          [0]
            bool bSafePoint
            ifItem iIfItem
              [0]
                bool bANDOR[2]
                num nSigIndex[3]
                num nSigType[3]
                num nValue[3]
            mdesc mMdesc
            num nActionIndex = 42
            num nDelay
            num nMoveType = 1
            num nPercentage
            num nSigValue = 1
        pointRx pPointRx[2] = {x=-245.0810672, y=-321.451661, z=639.817242, rx=-2.232299, ry=1.28487, rz=0.967617, shoulder=lefty, elbow=enegative, wrist=wpositive}
        string sID
      [8]
        bool bMarked
        jointRx jJointRx = {j1=-122.510061, j2=129.763772, j3=-115.645271, j4=180.40219, j5=16.691098, j6=-56.935013}
        pointRx pInter
        paraItem pParaItem
          [0]
            bool bSafePoint
            ifItem iIfItem
              [0]
                bool bANDOR[2]
                num nSigIndex[3]
                num nSigType[3]
                num nValue[3]
            mdesc mMdesc
            num nActionIndex = 42
            num nDelay
            num nMoveType = 1
            num nPercentage
            num nSigValue = 1
        pointRx pPointRx[2] = {x=-204.794752, y=-412.495541, z=639.817259, rx=-2.23161, ry=1.284656, rz=0.967787, shoulder=lefty, elbow=enegative, wrist=wpositive}
        string sID
      [9]
        bool bMarked
        jointRx jJointRx = {j1=-115.509708, j2=123.384757, j3=-95.0786351, j4=179.613978, j5=30.87235, j6=-63.211859}
        pointRx pInter
        paraItem pParaItem
          [0]
            bool bSafePoint
            ifItem iIfItem
              [0]
                bool bANDOR[2]
                num nSigIndex[3]
                num nSigType[3]
                num nValue[3]
            mdesc mMdesc
            num nActionIndex = 42
            num nDelay
            num nMoveType = 1
            num nPercentage
            num nSigValue = 1
        pointRx pPointRx[2] = {x=-204.829932, y=-549.361149, z=639.817236, rx=-2.230566, ry=1.283434, rz=0.967655, shoulder=lefty, elbow=enegative, wrist=wpositive}
        string sID
      [10]
        bool bMarked
        jointRx jJointRx = {j1=-115.168839, j2=115.765951, j3=-75.660997, j4=179.549971, j5=42.662693, j6=-65.612389}
        pointRx pInter
        paraItem pParaItem
          [0]
            bool bSafePoint
            ifItem iIfItem
              [0]
                bool bANDOR[2]
                num nSigIndex[3]
                num nSigType[3]
                num nValue[3]
            mdesc mMdesc
            num nActionIndex = 42
            num nDelay
            num nMoveType = 1
            num nPercentage
            num nSigValue = 1
        pointRx pPointRx[2] = {x=-243.328707, y=-641.656144, z=639.817272, rx=-2.184752, ry=1.363169, rz=-1.0929741, shoulder=lefty, elbow=enegative, wrist=wpositive}
        string sID
      [11]
        bool bMarked
        jointRx jJointRx = {j1=-103.18234, j2=119.0666826, j3=-83.752693, j4=178.724024, j5=37.773968, j6=-75.789236}
        pointRx pInter
        paraItem pParaItem
          [0]
            bool bSafePoint
            ifItem iIfItem
              [0]
                bool bANDOR[2]
                num nSigIndex[3]
                num nSigType[3]
                num nValue[3]
            mdesc mMdesc
            num nActionIndex = 42
            num nDelay
            num nMoveType = 1
            num nPercentage
            num nSigValue = 1
        pointRx pPointRx[2] = {x=-91.940597, y=-641.690605, z=639.817264, rx=-2.210413, ry=1.320263, rz=0.0285249, shoulder=lefty, elbow=enegative, wrist=wpositive}
        string sID
      [12]
        bool bMarked
        jointRx jJointRx = {j1=-96.605755, j2=119.651273, j3=-85.228552, j4=178.232883, j5=36.783421, j6=-81.95314}
        pointRx pInter
        paraItem pParaItem
          [0]
            bool bSafePoint
            ifItem iIfItem
              [0]
                bool bANDOR[2]
                num nSigIndex[3]
                num nSigType[3]
                num nValue[3]
            mdesc mMdesc
            num nActionIndex = 42
            num nDelay
            num nMoveType = 1
            num nPercentage
            num nSigValue = 1
        pointRx pPointRx[2] = {x=-14.68309, y=-641.690595, z=639.817262, rx=-2.210425, ry=1.321003, rz=0.029458, shoulder=lefty, elbow=enegative, wrist=wpositive}
        string sID
      [13]
        bool bMarked
        jointRx jJointRx = {j1=-101.415655, j2=125.744666, j3=-101.857376, j4=178.0690532, j5=26.328772, j6=-76.831785}
        pointRx pInter
        paraItem pParaItem
          [0]
            bool bSafePoint
            ifItem iIfItem
              [0]
                bool bANDOR[2]
                num nSigIndex[3]
                num nSigType[3]
                num nValue[3]
            mdesc mMdesc
            num nActionIndex = 42
            num nDelay
            num nMoveType = 1
            num nPercentage
            num nSigValue = 1
        pointRx pPointRx[2] = {x=-51.703517, y=-546.433248, z=639.817258, rx=-2.211187, ry=1.319905, rz=0.0291157, shoulder=lefty, elbow=enegative, wrist=wpositive}
        string sID
      [14]
        bool bMarked
        jointRx jJointRx = {j1=-104.908394, j2=131.188615, j3=-122.570612, j4=176.33465, j5=11.11624, j6=-71.475976}
        pointRx pInter
        paraItem pParaItem
          [0]
            bool bSafePoint
            ifItem iIfItem
              [0]
                bool bANDOR[2]
                num nSigIndex[3]
                num nSigType[3]
                num nValue[3]
            mdesc mMdesc
            num nActionIndex = 42
            num nDelay
            num nMoveType = 1
            num nPercentage
            num nSigValue = 1
        pointRx pPointRx[2] = {x=-51.703514, y=-412.500595, z=639.817231, rx=-2.211237, ry=1.319324, rz=0.0290677, shoulder=lefty, elbow=enegative, wrist=wpositive}
        string sID
      [15]
        bool bMarked
        jointRx jJointRx = {j1=-113.792229, j2=132.0385925, j3=-133.203423, j4=167.238796, j5=1.425916, j6=-53.439675}
        pointRx pInter
        paraItem pParaItem
          [0]
            bool bSafePoint
            ifItem iIfItem
              [0]
                bool bANDOR[2]
                num nSigIndex[3]
                num nSigType[3]
                num nValue[3]
            mdesc mMdesc
            num nActionIndex = 42
            num nDelay
            num nMoveType = 1
            num nPercentage
            num nSigValue = 1
        pointRx pPointRx[2] = {x=-86.764293, y=-327.545777, z=639.814183, rx=-2.211628, ry=1.318889, rz=0.029149, shoulder=lefty, elbow=enegative, wrist=wpositive}
        string sID
      [16]
        bool bMarked
        jointRx jJointRx = {j1=-111.801102, j2=131.0492813, j3=-121.763212, j4=165.182491, j5=10.00939302, j6=-125.703677}
        pointRx pInter
        paraItem pParaItem
          [0]
            bool bSafePoint
            ifItem iIfItem
              [0]
                bool bANDOR[2]
                num nSigIndex[3]
                num nSigType[3]
                num nValue[3]
            mdesc mMdesc
            num nActionIndex = 42
            num nDelay
            num nMoveType = 1
            num nPercentage
            num nSigValue = 1
        pointRx pPointRx[2] = {x=-94.727754, y=-431.297828, z=639.823313, rx=0.578297, ry=2.512713, rz=-72.12797, shoulder=lefty, elbow=enegative, wrist=wpositive}
        string sID
      [17]
        bool bMarked
        jointRx jJointRx = {j1=-100.696291, j2=131.394596, j3=-123.887641, j4=160.749292, j5=7.838779, j6=-132.328285}
        pointRx pInter
        paraItem pParaItem
          [0]
            bool bSafePoint
            ifItem iIfItem
              [0]
                bool bANDOR[2]
                num nSigIndex[3]
                num nSigType[3]
                num nValue[3]
            mdesc mMdesc
            num nActionIndex = 42
            num nDelay
            num nMoveType = 1
            num nPercentage
            num nSigValue = 1
        pointRx pPointRx[2] = {x=-7.700551, y=-431.29776, z=639.823315, rx=0.578366, ry=2.513634, rz=-72.118873, shoulder=lefty, elbow=enegative, wrist=wpositive}
        string sID
      [18]
        bool bMarked
        jointRx jJointRx = {j1=-85.175274, j2=131.219929, j3=-122.767363, j4=172.20701, j5=10.687341, j6=-85.487938}
        pointRx pInter
        paraItem pParaItem
          [0]
            bool bSafePoint
            ifItem iIfItem
              [0]
                bool bANDOR[2]
                num nSigIndex[3]
                num nSigType[3]
                num nValue[3]
            mdesc mMdesc
            num nActionIndex = 42
            num nDelay
            num nMoveType = 1
            num nPercentage
            num nSigValue = 1
        pointRx pPointRx[2] = {x=97.129831, y=-406.771802, z=639.823216, rx=-2.251869, ry=1.255999, rz=1.675152, shoulder=lefty, elbow=enegative, wrist=wpositive}
        string sID
      [19]
        bool bMarked
        jointRx jJointRx = {j1=-78.327634, j2=132.0275027, j3=-133.511556, j4=105.524405, j5=1.749155, j6=-25.524463}
        pointRx pInter
        paraItem pParaItem
          [0]
            bool bSafePoint
            ifItem iIfItem
              [0]
                bool bANDOR[2]
                num nSigIndex[3]
                num nSigType[3]
                num nValue[3]
            mdesc mMdesc
            num nActionIndex = 42
            num nDelay
            num nMoveType
            num nPercentage
            num nSigValue = 1
        pointRx pPointRx[2] = {x=131.681956, y=-317.592689, z=639.818955, rx=-2.252815, ry=1.25559, rz=1.675166, shoulder=lefty, elbow=enegative, wrist=wpositive}
        string sID
      [20]
        bool bMarked
        jointRx jJointRx = {j1=-86.344906, j2=125.635703, j3=-101.533058, j4=176.84641, j5=26.303372, j6=-89.150638}
        pointRx pInter
        paraItem pParaItem
          [0]
            bool bSafePoint
            ifItem iIfItem
              [0]
                bool bANDOR[2]
                num nSigIndex[3]
                num nSigType[3]
                num nValue[3]
            mdesc mMdesc
            num nActionIndex = 42
            num nDelay
            num nMoveType = 1
            num nPercentage
            num nSigValue = 1
        pointRx pPointRx[2] = {x=97.129791, y=-544.994507, z=639.823164, rx=-2.250847, ry=1.25596, rz=1.67509, shoulder=lefty, elbow=enegative, wrist=wpositive}
        string sID
      [21]
        bool bMarked
        jointRx jJointRx = {j1=-90.472886, j2=120.653514, j3=-87.796909, j4=177.850277, j5=35.136858, j6=-86.0941041}
        pointRx pInter
        paraItem pParaItem
          [0]
            bool bSafePoint
            ifItem iIfItem
              [0]
                bool bANDOR[2]
                num nSigIndex[3]
                num nSigType[3]
                num nValue[3]
            mdesc mMdesc
            num nActionIndex = 42
            num nDelay
            num nMoveType = 1
            num nPercentage
            num nSigValue = 1
        pointRx pPointRx[2] = {x=55.621844, y=-626.948778, z=639.823217, rx=-2.25099, ry=1.255655, rz=1.674992, shoulder=lefty, elbow=enegative, wrist=wpositive}
        string sID
      [22]
        bool bMarked
        jointRx jJointRx = {j1=-83.248503, j2=126.765701, j3=-105.0119337, j4=185.0332952, j5=23.463189, j6=-12.861735}
        pointRx pInter
        paraItem pParaItem
          [0]
            bool bSafePoint
            ifItem iIfItem
              [0]
                bool bANDOR[2]
                num nSigIndex[3]
                num nSigType[3]
                num nValue[3]
            mdesc mMdesc
            num nActionIndex = 42
            num nDelay
            num nMoveType = 1
            num nPercentage
            num nSigValue = 1
        pointRx pPointRx[2] = {x=95.0604108, y=-526.24744, z=639.845413, rx=-1.382011, ry=-2.179455, rz=88.510933, shoulder=lefty, elbow=enegative, wrist=wpositive}
        string sID
      [23]
        bool bMarked
        jointRx jJointRx = {j1=-102.947247, j2=123.371825, j3=-104.720974, j4=140.865912, j5=30.580144, j6=47.745938}
        pointRx pInter
        paraItem pParaItem
          [0]
            bool bSafePoint
            ifItem iIfItem
              [0]
                bool bANDOR[2]
                num nSigIndex[3]
                num nSigType[3]
                num nValue[3]
            mdesc mMdesc
            num nActionIndex = 42
            num nDelay
            num nMoveType = 1
            num nPercentage
            num nSigValue = 1
        pointRx pPointRx[2] = {x=95.0560257, y=-526.230668, z=639.854281, rx=-1.467206, ry=19.573094, rz=89.0544323, shoulder=lefty, elbow=enegative, wrist=wpositive}
        string sID
      [24]
        bool bMarked
        jointRx jJointRx = {j1=-105.42444, j2=126.319202, j3=-118.0699052, j4=127.900909, j5=23.640583, j6=64.972841}
        pointRx pInter
        paraItem pParaItem
          [0]
            bool bSafePoint
            ifItem iIfItem
              [0]
                bool bANDOR[2]
                num nSigIndex[3]
                num nSigType[3]
                num nValue[3]
            mdesc mMdesc
            num nActionIndex = 42
            num nDelay
            num nMoveType = 1
            num nPercentage
            num nSigValue = 1
        pointRx pPointRx[2] = {x=95.0558629, y=-438.311234, z=639.854334, rx=-1.468101, ry=19.566479, rz=89.0544973, shoulder=lefty, elbow=enegative, wrist=wpositive}
        string sID
      [25]
        bool bMarked
        jointRx jJointRx = {j1=-112.0262192, j2=125.853254, j3=-136.407591, j4=84.864182, j5=17.615577, j6=117.594482}
        pointRx pInter
        paraItem pParaItem
          [0]
            bool bSafePoint
            ifItem iIfItem
              [0]
                bool bANDOR[2]
                num nSigIndex[3]
                num nSigType[3]
                num nValue[3]
            mdesc mMdesc
            num nActionIndex = 42
            num nDelay
            num nMoveType = 1
            num nPercentage
            num nSigValue = 1
        pointRx pPointRx[2] = {x=95.0562279, y=-300.211931, z=639.855152, rx=-1.466155, ry=19.566406, rz=89.0540412, shoulder=lefty, elbow=enegative, wrist=wpositive}
        string sID
      [26]
        bool bMarked
        jointRx jJointRx = {j1=-98.853409, j2=130.526556, j3=-129.84131, j4=190.937055, j5=1.850619, j6=112.778311}
        pointRx pInter
        paraItem pParaItem
          [0]
            bool bSafePoint
            ifItem iIfItem
              [0]
                bool bANDOR[2]
                num nSigIndex[3]
                num nSigType[3]
                num nValue[3]
            mdesc mMdesc
            num nActionIndex = 42
            num nDelay
            num nMoveType = 1
            num nPercentage
            num nSigValue = 1
        pointRx pPointRx[2] = {x=-10.299262, y=-371.0877835, z=648.6975, rx=-1.172321, ry=-0.172701, rz=-155.141909, shoulder=lefty, elbow=enegative, wrist=wpositive}
        string sID
      [27]
        bool bMarked
        jointRx jJointRx = {j1=-87.556691, j2=130.508226, j3=-129.0706324, j4=182.704505, j5=2.618876, j6=109.713672}
        pointRx pInter
        paraItem pParaItem
          [0]
            bool bSafePoint
            ifItem iIfItem
              [0]
                bool bANDOR[2]
                num nSigIndex[3]
                num nSigType[3]
                num nValue[3]
            mdesc mMdesc
            num nActionIndex = 42
            num nDelay
            num nMoveType = 1
            num nPercentage
            num nSigValue = 1
        pointRx pPointRx[2] = {x=64.800708, y=-371.087733, z=648.697509, rx=-1.172034, ry=-0.173648, rz=-155.14184, shoulder=lefty, elbow=enegative, wrist=wpositive}
        string sID
      [28]
        bool bMarked
        jointRx jJointRx = {j1=-76.56227, j2=130.441663, j3=-127.63649, j4=178.503737, j5=3.987538, j6=102.915897}
        pointRx pInter
        paraItem pParaItem
          [0]
            bool bSafePoint
            ifItem iIfItem
              [0]
                bool bANDOR[2]
                num nSigIndex[3]
                num nSigType[3]
                num nValue[3]
            mdesc mMdesc
            num nActionIndex = 42
            num nDelay
            num nMoveType = 1
            num nPercentage
            num nSigValue = 1
        pointRx pPointRx[2] = {x=138.739125, y=-361.605648, z=648.697463, rx=-1.172859, ry=-0.173244, rz=-155.141862, shoulder=lefty, elbow=enegative, wrist=wpositive}
        string sID
      [29]
        bool bMarked
        jointRx jJointRx = {j1=-65.258595, j2=131.722388, j3=-131.258412, j4=149.998176, j5=1.563572, j6=95.282187}
        pointRx pInter
        paraItem pParaItem
          [0]
            bool bSafePoint
            ifItem iIfItem
              [0]
                bool bANDOR[2]
                num nSigIndex[3]
                num nSigType[3]
                num nValue[3]
            mdesc mMdesc
            num nActionIndex = 42
            num nDelay
            num nMoveType = 1
            num nPercentage
            num nSigValue = 1
        pointRx pPointRx[2] = {x=203.481922, y=-305.793086, z=642.0323173, rx=-1.135624, ry=0.337465, rz=-179.971722, shoulder=lefty, elbow=enegative, wrist=wpositive}
        string sID
      [30]
        bool bMarked
        jointRx jJointRx = {j1=-75.287181, j2=130.366871, j3=-119.512671, j4=177.0231421, j5=11.88329, j6=78.230615}
        pointRx pInter
        paraItem pParaItem
          [0]
            bool bSafePoint
            ifItem iIfItem
              [0]
                bool bANDOR[2]
                num nSigIndex[3]
                num nSigType[3]
                num nValue[3]
            mdesc mMdesc
            num nActionIndex = 42
            num nDelay
            num nMoveType = 1
            num nPercentage
            num nSigValue = 1
        pointRx pPointRx[2] = {x=166.551107, y=-416.353492, z=642.0259775, rx=-1.135878, ry=0.33525, rz=-179.971835, shoulder=lefty, elbow=enegative, wrist=wpositive}
        string sID
      [31]
        bool bMarked
        jointRx jJointRx = {j1=-78.750875, j2=124.345332, j3=-98.32121, j4=178.789895, j5=27.0774003, j6=79.858309}
        pointRx pInter
        paraItem pParaItem
          [0]
            bool bSafePoint
            ifItem iIfItem
              [0]
                bool bANDOR[2]
                num nSigIndex[3]
                num nSigType[3]
                num nValue[3]
            mdesc mMdesc
            num nActionIndex = 42
            num nDelay
            num nMoveType = 1
            num nPercentage
            num nSigValue = 1
        pointRx pPointRx[2] = {x=166.551118, y=-556.425136, z=642.0259681, rx=-1.135398, ry=0.335774, rz=-179.971779, shoulder=lefty, elbow=enegative, wrist=wpositive}
        string sID
      [32]
        bool bMarked
        jointRx jJointRx = {j1=-83.872725, j2=117.4103, j3=-80.0479523, j4=179.268733, j5=38.458687, j6=84.472525}
        pointRx pInter
        paraItem pParaItem
          [0]
            bool bSafePoint
            ifItem iIfItem
              [0]
                bool bANDOR[2]
                num nSigIndex[3]
                num nSigType[3]
                num nValue[3]
            mdesc mMdesc
            num nActionIndex = 42
            num nDelay
            num nMoveType = 1
            num nPercentage
            num nSigValue = 1
        pointRx pPointRx[2] = {x=125.777964, y=-666.0321845, z=642.0361412, rx=-1.136355, ry=0.335436, rz=-179.973852, shoulder=lefty, elbow=enegative, wrist=wpositive}
        string sID
      [33]
        bool bMarked
        jointRx jJointRx = {j1=-78.0158878, j2=116.00480506, j3=-76.619863, j4=179.128646, j5=40.428713, j6=78.707523}
        pointRx pInter
        paraItem pParaItem
          [0]
            bool bSafePoint
            ifItem iIfItem
              [0]
                bool bANDOR[2]
                num nSigIndex[3]
                num nSigType[3]
                num nValue[3]
            mdesc mMdesc
            num nActionIndex = 42
            num nDelay
            num nMoveType = 1
            num nPercentage
            num nSigValue = 1
        pointRx pPointRx[2] = {x=197.538696, y=-666.0666154, z=642.0361247, rx=-1.135138, ry=0.336712, rz=-179.973468, shoulder=lefty, elbow=enegative, wrist=wpositive}
        string sID
      [34]
        bool bMarked
        jointRx jJointRx = {j1=-72.0822941, j2=113.707363, j3=-71.14889, j4=179.0271553, j5=43.540761, j6=72.816847}
        pointRx pInter
        paraItem pParaItem
          [0]
            bool bSafePoint
            ifItem iIfItem
              [0]
                bool bANDOR[2]
                num nSigIndex[3]
                num nSigType[3]
                num nValue[3]
            mdesc mMdesc
            num nActionIndex = 42
            num nDelay
            num nMoveType = 1
            num nPercentage
            num nSigValue = 1
        pointRx pPointRx[2] = {x=274.0463743, y=-666.0377191, z=642.0648113, rx=-1.136874, ry=0.336734, rz=-179.973059, shoulder=lefty, elbow=enegative, wrist=wpositive}
        string sID
      [35]
        bool bMarked
        jointRx jJointRx = {j1=-68.231832, j2=114.0101375, j3=-71.862732, j4=178.925387, j5=43.085151, j6=69.0461931}
        pointRx pInter
        paraItem pParaItem
          [0]
            bool bSafePoint
            ifItem iIfItem
              [0]
                bool bANDOR[2]
                num nSigIndex[3]
                num nSigType[3]
                num nValue[3]
            mdesc mMdesc
            num nActionIndex = 42
            num nDelay
            num nMoveType = 1
            num nPercentage
            num nSigValue = 1
        pointRx pPointRx[2] = {x=317.646205, y=-643.356636, z=642.0648372, rx=-1.138401, ry=0.335813, rz=-179.973153, shoulder=lefty, elbow=enegative, wrist=wpositive}
        string sID
      [36]
        bool bMarked
        jointRx jJointRx = {j1=-65.210051, j2=120.724606, j3=-88.443145, j4=178.570875, j5=33.182263, j6=66.435792}
        pointRx pInter
        paraItem pParaItem
          [0]
            bool bSafePoint
            ifItem iIfItem
              [0]
                bool bANDOR[2]
                num nSigIndex[3]
                num nSigType[3]
                num nValue[3]
            mdesc mMdesc
            num nActionIndex = 42
            num nDelay
            num nMoveType = 1
            num nPercentage
            num nSigValue = 1
        pointRx pPointRx[2] = {x=317.646188, y=-552.240414, z=642.0648293, rx=-1.138291, ry=0.335792, rz=-179.973173, shoulder=lefty, elbow=enegative, wrist=wpositive}
        string sID
      [37]
        bool bMarked
        jointRx jJointRx = {j1=-59.269672, j2=127.333625, j3=-107.550013, j4=177.526605, j5=20.607904, j6=61.614613}
        pointRx pInter
        paraItem pParaItem
          [0]
            bool bSafePoint
            ifItem iIfItem
              [0]
                bool bANDOR[2]
                num nSigIndex[3]
                num nSigType[3]
                num nValue[3]
            mdesc mMdesc
            num nActionIndex = 42
            num nDelay
            num nMoveType = 1
            num nPercentage
            num nSigValue = 1
        pointRx pPointRx[2] = {x=317.646169, y=-421.622338, z=642.0648205, rx=-1.138138, ry=0.335927, rz=-179.973153, shoulder=lefty, elbow=enegative, wrist=wpositive}
        string sID
      [38]
        bool bMarked
        jointRx jJointRx = {j1=-56.529834, j2=131.219574, j3=-124.66737, j4=172.915754, j5=7.371604, j6=63.585523}
        pointRx pInter
        paraItem pParaItem
          [0]
            bool bSafePoint
            ifItem iIfItem
              [0]
                bool bANDOR[2]
                num nSigIndex[3]
                num nSigType[3]
                num nValue[3]
            mdesc mMdesc
            num nActionIndex = 42
            num nDelay
            num nMoveType = 1
            num nPercentage
            num nSigValue = 1
        pointRx pPointRx[2] = {x=275.258961, y=-311.334534, z=642.0647626, rx=-1.137088, ry=0.335146, rz=-179.97331, shoulder=lefty, elbow=enegative, wrist=wpositive}
        string sID
      [39]
        bool bMarked
        jointRx jJointRx = {j1=-63.306074, j2=128.457716, j3=-111.487898, j4=177.354165, j5=17.85182, j6=65.854127}
        pointRx pInter
        paraItem pParaItem
          [0]
            bool bSafePoint
            ifItem iIfItem
              [0]
                bool bANDOR[2]
                num nSigIndex[3]
                num nSigType[3]
                num nValue[3]
            mdesc mMdesc
            num nActionIndex = 42
            num nDelay
            num nMoveType = 1
            num nPercentage
            num nSigValue = 1
        pointRx pPointRx[2] = {x=275.293372, y=-420.450747, z=642.0648054, rx=-1.136295, ry=0.336239, rz=-179.973341, shoulder=lefty, elbow=enegative, wrist=wpositive}
        string sID
      [40]
        bool bMarked
        jointRx jJointRx = {j1=-81.00112581, j2=130.644686, j3=-121.00772478, j4=177.263665, j5=10.719901, j6=83.717831}
        pointRx pInter
        paraItem pParaItem
          [0]
            bool bSafePoint
            ifItem iIfItem
              [0]
                bool bANDOR[2]
                num nSigIndex[3]
                num nSigType[3]
                num nValue[3]
            mdesc mMdesc
            num nActionIndex = 42
            num nDelay
            num nMoveType = 1
            num nPercentage
            num nSigValue = 1
        pointRx pPointRx[2] = {x=121.697258, y=-420.415642, z=642.064816, rx=-1.13739, ry=0.335022, rz=-179.973377, shoulder=lefty, elbow=enegative, wrist=wpositive}
        string sID
      [41]
        bool bMarked
        jointRx jJointRx = {j1=-101.57564, j2=130.996968, j3=-123.11763, j4=179.378674, j5=9.0641696, j6=102.209948}
        pointRx pInter
        paraItem pParaItem
          [0]
            bool bSafePoint
            ifItem iIfItem
              [0]
                bool bANDOR[2]
                num nSigIndex[3]
                num nSigType[3]
                num nValue[3]
            mdesc mMdesc
            num nActionIndex = 42
            num nDelay
            num nMoveType = 1
            num nPercentage
            num nSigValue = 1
        pointRx pPointRx[2] = {x=-34.195927, y=-420.382673, z=642.0719086, rx=-1.140588, ry=0.333521, rz=-179.976951, shoulder=lefty, elbow=enegative, wrist=wpositive}
        string sID
      [42]
        bool bMarked
        jointRx jJointRx = {j1=-117.910926, j2=130.159863, j3=-118.527747, j4=181.0779949, j5=12.798502, j6=116.877037}
        pointRx pInter
        paraItem pParaItem
          [0]
            bool bSafePoint
            ifItem iIfItem
              [0]
                bool bANDOR[2]
                num nSigIndex[3]
                num nSigType[3]
                num nValue[3]
            mdesc mMdesc
            num nActionIndex = 42
            num nDelay
            num nMoveType = 1
            num nPercentage
            num nSigValue = 1
        pointRx pPointRx[2] = {x=-168.460127, y=-420.382669, z=642.071906, rx=-1.140562, ry=0.333907, rz=-179.976921, shoulder=lefty, elbow=enegative, wrist=wpositive}
        string sID
      [43]
        bool bMarked
        jointRx jJointRx = {j1=-132.269491, j2=127.123938, j3=-106.855674, j4=181.429188, j5=21.342688, j6=130.953129}
        pointRx pInter
        paraItem pParaItem
          [0]
            bool bSafePoint
            ifItem iIfItem
              [0]
                bool bANDOR[2]
                num nSigIndex[3]
                num nSigType[3]
                num nValue[3]
            mdesc mMdesc
            num nActionIndex = 42
            num nDelay
            num nMoveType = 1
            num nPercentage
            num nSigValue = 1
        pointRx pPointRx[2] = {x=-320.674662, y=-420.382638, z=642.0718966, rx=-1.140431, ry=0.333681, rz=-179.976981, shoulder=lefty, elbow=enegative, wrist=wpositive}
        string sID
      [44]
        bool bMarked
        jointRx jJointRx = {j1=-142.441106, j2=120.824327, j3=-88.705493, j4=181.282913, j5=33.0850501, j6=141.380041}
        pointRx pInter
        paraItem pParaItem
          [0]
            bool bSafePoint
            ifItem iIfItem
              [0]
                bool bANDOR[2]
                num nSigIndex[3]
                num nSigType[3]
                num nValue[3]
            mdesc mMdesc
            num nActionIndex = 42
            num nDelay
            num nMoveType = 1
            num nPercentage
            num nSigValue = 1
        pointRx pPointRx[2] = {x=-474.689621, y=-420.382631, z=642.0718894, rx=-1.140119, ry=0.333784, rz=-179.976923, shoulder=lefty, elbow=enegative, wrist=wpositive}
        string sID
      [45]
        bool bMarked
        jointRx jJointRx = {j1=-138.108258, j2=121.207146, j3=-89.710766, j4=181.162609, j5=32.51161, j6=137.142341}
        pointRx pInter
        paraItem pParaItem
          [0]
            bool bSafePoint
            ifItem iIfItem
              [0]
                bool bANDOR[2]
                num nSigIndex[3]
                num nSigType[3]
                num nValue[3]
            mdesc mMdesc
            num nActionIndex = 42
            num nDelay
            num nMoveType = 1
            num nPercentage
            num nSigValue = 1
        pointRx pPointRx[2] = {x=-436.796862, y=-451.644484, z=642.07189, rx=-1.139469, ry=0.334472, rz=-179.976638, shoulder=lefty, elbow=enegative, wrist=wpositive}
        string sID
      [46]
        bool bMarked
        jointRx jJointRx = {j1=-127.70596, j2=126.693595, j3=-105.454305, j4=181.135682, j5=22.350888, j6=126.671469}
        pointRx pInter
        paraItem pParaItem
          [0]
            bool bSafePoint
            ifItem iIfItem
              [0]
                bool bANDOR[2]
                num nSigIndex[3]
                num nSigType[3]
                num nValue[3]
            mdesc mMdesc
            num nActionIndex = 42
            num nDelay
            num nMoveType = 1
            num nPercentage
            num nSigValue = 1
        pointRx pPointRx[2] = {x=-290.683508, y=-451.609469, z=642.07191, rx=-1.140457, ry=0.335724, rz=-179.976594, shoulder=lefty, elbow=enegative, wrist=wpositive}
        string sID
      [47]
        bool bMarked
        jointRx jJointRx = {j1=-77.238254, j2=129.340507, j3=-114.913945, j4=177.831104, j5=15.475362, j6=79.35375}
        pointRx pInter
        paraItem pParaItem
          [0]
            bool bSafePoint
            ifItem iIfItem
              [0]
                bool bANDOR[2]
                num nSigIndex[3]
                num nSigType[3]
                num nValue[3]
            mdesc mMdesc
            num nActionIndex = 42
            num nDelay
            num nMoveType = 1
            num nPercentage
            num nSigValue = 1
        pointRx pPointRx[2] = {x=158.729452, y=-451.609464, z=642.0719065, rx=-1.140389, ry=0.334964, rz=-179.976748, shoulder=lefty, elbow=enegative, wrist=wpositive}
        string sID
      [48]
        bool bMarked
        jointRx jJointRx = {j1=-63.488687, j2=124.208026, j3=-97.940675, j4=178.228458, j5=27.14867, j6=65.0910716}
        pointRx pInter
        paraItem pParaItem
          [0]
            bool bSafePoint
            ifItem iIfItem
              [0]
                bool bANDOR[2]
                num nSigIndex[3]
                num nSigType[3]
                num nValue[3]
            mdesc mMdesc
            num nActionIndex = 42
            num nDelay
            num nMoveType = 1
            num nPercentage
            num nSigValue = 1
        pointRx pPointRx[2] = {x=310.830797, y=-495.30753, z=642.0718875, rx=-1.139453, ry=0.33486, rz=-179.976891, shoulder=lefty, elbow=enegative, wrist=wpositive}
        string sID
      [49]
        bool bMarked
        jointRx jJointRx = {j1=-78.0579912, j2=127.559769, j3=-108.316642, j4=178.378161, j5=20.297351, j6=79.604006}
        pointRx pInter
        paraItem pParaItem
          [0]
            bool bSafePoint
            ifItem iIfItem
              [0]
                bool bANDOR[2]
                num nSigIndex[3]
                num nSigType[3]
                num nValue[3]
            mdesc mMdesc
            num nActionIndex = 42
            num nDelay
            num nMoveType = 1
            num nPercentage
            num nSigValue = 1
        pointRx pPointRx[2] = {x=160.873249, y=-495.272541, z=642.0719096, rx=-1.140489, ry=0.333782, rz=-179.976981, shoulder=lefty, elbow=enegative, wrist=wpositive}
        string sID
      [50]
        bool bMarked
        jointRx jJointRx = {j1=-83.970136, j2=129.00855342, j3=-113.590578, j4=181.751291, j5=14.32041, j6=-96.622719}
        pointRx pInter
        paraItem pParaItem
          [0]
            bool bSafePoint
            ifItem iIfItem
              [0]
                bool bANDOR[2]
                num nSigIndex[3]
                num nSigType[3]
                num nValue[3]
            mdesc mMdesc
            num nActionIndex = 42
            num nDelay
            num nMoveType = 1
            num nPercentage
            num nSigValue = 1
        pointRx pPointRx[2] = {x=98.789636, y=-495.232609, z=642.0875542, rx=1.143362, ry=-0.31475, rz=1.103019, shoulder=lefty, elbow=enegative, wrist=wpositive}
        string sID
      [51]
        bool bMarked
        jointRx jJointRx = {j1=-101.251443, j2=129.329307, j3=-114.876217, j4=180.377122, j5=13.270505, j6=-78.0149862}
        pointRx pInter
        paraItem pParaItem
          [0]
            bool bSafePoint
            ifItem iIfItem
              [0]
                bool bANDOR[2]
                num nSigIndex[3]
                num nSigType[3]
                num nValue[3]
            mdesc mMdesc
            num nActionIndex = 42
            num nDelay
            num nMoveType = 1
            num nPercentage
            num nSigValue = 1
        pointRx pPointRx[2] = {x=-48.311282, y=-495.232554, z=642.0875543, rx=1.143247, ry=-0.315683, rz=1.102879, shoulder=lefty, elbow=enegative, wrist=wpositive}
        string sID
      [52]
        bool bMarked
        jointRx jJointRx = {j1=-117.974593, j2=127.746571, j3=-108.963712, j4=179.150072, j5=17.626951, j6=-60.118292}
        pointRx pInter
        paraItem pParaItem
          [0]
            bool bSafePoint
            ifItem iIfItem
              [0]
                bool bANDOR[2]
                num nSigIndex[3]
                num nSigType[3]
                num nValue[3]
            mdesc mMdesc
            num nActionIndex = 42
            num nDelay
            num nMoveType = 1
            num nPercentage
            num nSigValue = 1
        pointRx pPointRx[2] = {x=-203.879984, y=-495.232578, z=642.0875477, rx=1.143192, ry=-0.315734, rz=1.102838, shoulder=lefty, elbow=enegative, wrist=wpositive}
        string sID
      [53]
        bool bMarked
        jointRx jJointRx = {j1=-130.30363, j2=123.943868, j3=-97.190977, j4=178.849142, j5=25.681002, j6=-47.564193}
        pointRx pInter
        paraItem pParaItem
          [0]
